DATA_BLOCK "GDB_OperationsTest"
{ S7_Optimized_Access := 'TRUE' }
VERSION : 0.1
NON_RETAIN
"FB_OperationsTest"
BEGIN
END_DATA_BLOCK
